(* IEC 61131-3 sources: SRCI_CLIENT_PLC/RobotLibrary/Library/Structures/Telegram, 1 file *)

(* ---- Telegram.st ---- *)
{attribute 'pack_mode' := '1'}
// -------------------------------------------------------------------------
//  SRCI Robot Library
// -------------------------------------------------------------------------
//
//  Object:      Telegram
//  Author:      Thorsten Brach
//  Date:        2024-06-01
//
//  Description:
//
//
//  Copyright:
//    (C) 2024 Thorsten Brach. All rights reserved
//             Licensed under the MIT License.
//
//  Disclaimer:
//    This project is provided without any guarantee and can be used for
//    private and commercial purposes. Any use is at the user’s
//    own risk and responsibility.
//
// -------------------------------------------------------------------------
TYPE Telegram :
STRUCT
  /// PLC to Robot
  PlcToRob : TelegramPlcToRob;
  /// Robot to PLC
  RobToPlc : TelegramRobToPlc;
END_STRUCT
END_TYPE
